{attribute 'linkalways'}
{attribute 'no_explicit_call' := 'This FB is a CLASS and must be accessed using methods or properties'}
{attribute 'enable_dynamic_creation'}
FUNCTION_BLOCK Node_F_VN_ReshapeImage EXTENDS VisionNode
VAR
    ipSrcImage : _ITcVnImage;
    ipDestImage : _ITcVnImage;
    aNewShape : _TcVnArray33_UDINT;
    hrPrev : _HRESULT(S_OK);
    hresult : _HRESULT(S_OK);
END_VAR

METHOD PUBLIC Clone : I_Node
VAR
    pNode : POINTER TO Node_F_VN_ReshapeImage;
END_VAR
pNode := __NEW(Node_F_VN_ReshapeImage);
Clone := pNode^;
END_METHOD

METHOD FB_init : BOOL
VAR_INPUT
    bInitRetains : BOOL;
    bInCopyCode : BOOL;
END_VAR
AddInput('ipSrcImage', ipSrcImage);
AddParameter('aNewShape', aNewShape);
AddInput('hrPrev', hrPrev);
AddOutput('ipDestImage', ipDestImage);
AddOutput('hresult', hresult);
END_METHOD

METHOD PROTECTED OnExecute
hresult.Value := F_VN_ReshapeImage(
    ipSrcImage := ipSrcImage.Value,
    ipDestImage := ipDestImage.Value,
    aNewShape := aNewShape.Value,
    hrPrev := hrPrev.Value);
END_METHOD

METHOD PUBLIC PreExecutionCheck
VAR_INPUT
    Check : I_PreExecutionChecks;
END_VAR
VAR
    i : UDINT;
    zeroDimensions : UDINT;
    dimensionCountIsValid : BOOL;
END_VAR
Check.IsTrue(ipSrcImage.IsValid, 'ipSrcImage must contain an image');
Check.IsTrue(ipSrcImage.HasChannelCount(1), 'ipSrcImage must have 1 channel');

dimensionCountIsValid := (aNewShape.Value[0] >= 1) AND (aNewShape.Value[0] <= 32);
Check.IsTrue(dimensionCountIsValid, 'aNewShape[0] must give the number of dimensions (1 to 32)');
IF dimensionCountIsValid THEN
    FOR i := 1 TO aNewShape.Value[0] DO
        IF aNewShape.Value[i] = 0 THEN
            zeroDimensions := zeroDimensions + 1;
        END_IF
    END_FOR
END_IF
Check.IsTrue(zeroDimensions <= 1, 'Only one dimension of aNewShape may be 0');
END_METHOD

END_FUNCTION_BLOCK

(* stored: Version 1.1.0.1, ProductVersion 3.1.4026.19
   POU Node_F_VN_ReshapeImage: Id {7b6180d5-e120-4fae-9d41-b75e99336d0c}, SpecialFunc None
   Folder Constructor: Id {a6cbb446-f233-4be4-ad67-a88d2891f0ed}
   Method Clone: Id {814c8aed-005a-470a-a7b7-0ab939f9b0f4}
   Method FB_init: Id {07bb4bb8-e143-4f01-b0ec-f21c4b8903a9}
   Method OnExecute: Id {dabfe9f2-900f-4049-9e40-d7ce007d4f44}
   Method PreExecutionCheck: Id {f926223b-47ea-4bbd-9021-94136e2bcd00} *)
